(* IEC 61131-3 sources: rusty/tests/lit/cfc/blocks/program_call, 2 files *)

(* ---- accumulator.st ---- *)
PROGRAM accumulator
VAR_INPUT
    step : DINT;
END_VAR
VAR_IN_OUT
    total : DINT;
END_VAR
VAR_OUTPUT
    doubled : DINT;
END_VAR
    total := total + step;
    doubled := total * 2;
END_PROGRAM

(* ---- main.st ---- *)
FUNCTION main : DINT
    program_call();
    program_call();
    // CHECK: total = 6, result = 12
    printf('total = %d, result = %d$N', program_call.runningTotal, program_call.result);
END_FUNCTION
